FUNCTION_BLOCK VALVE_MANIFOLD (* Migrated from IEC 61131-3 ST *)
  (* Standard: 61499-2 *)
  (* Version 1.0, 2026-11-06, st2fb *)
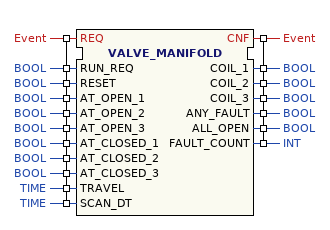
  EVENT_INPUT
    REQ WITH RUN_REQ, RESET, AT_OPEN_1, AT_OPEN_2, AT_OPEN_3, AT_CLOSED_1, AT_CLOSED_2, AT_CLOSED_3, TRAVEL, SCAN_DT;
  END_EVENT
  EVENT_OUTPUT
    CNF WITH COIL_1, COIL_2, COIL_3, ANY_FAULT, ALL_OPEN, FAULT_COUNT;
  END_EVENT
  VAR_INPUT
    RUN_REQ : BOOL;
    RESET : BOOL;
    AT_OPEN_1 : BOOL;
    AT_OPEN_2 : BOOL;
    AT_OPEN_3 : BOOL;
    AT_CLOSED_1 : BOOL;
    AT_CLOSED_2 : BOOL;
    AT_CLOSED_3 : BOOL;
    TRAVEL : TIME;
    SCAN_DT : TIME;
  END_VAR
  VAR_OUTPUT
    COIL_1 : BOOL;
    COIL_2 : BOOL;
    COIL_3 : BOOL;
    ANY_FAULT : BOOL;
    ALL_OPEN : BOOL;
    FAULT_COUNT : INT;
  END_VAR
  VAR
    ST2FB_NOW : TIME := T#0s;
    V1_OPEN_CMD : BOOL;
    V1_COIL : BOOL;
    V1_FAULT : BOOL;
    V1_OPENED : BOOL;
    V1_W_IN : BOOL;
    V1_W_PT : TIME;
    V1_W_Q : BOOL;
    V1_W_ET : TIME;
    V1_W_STATE : INT;
    V1_W_PREV_IN : BOOL;
    V1_W_START_TIME : TIME;
    V2_OPEN_CMD : BOOL;
    V2_COIL : BOOL;
    V2_FAULT : BOOL;
    V2_OPENED : BOOL;
    V2_W_IN : BOOL;
    V2_W_PT : TIME;
    V2_W_Q : BOOL;
    V2_W_ET : TIME;
    V2_W_STATE : INT;
    V2_W_PREV_IN : BOOL;
    V2_W_START_TIME : TIME;
    V3_OPEN_CMD : BOOL;
    V3_COIL : BOOL;
    V3_FAULT : BOOL;
    V3_OPENED : BOOL;
    V3_W_IN : BOOL;
    V3_W_PT : TIME;
    V3_W_Q : BOOL;
    V3_W_ET : TIME;
    V3_W_STATE : INT;
    V3_W_PREV_IN : BOOL;
    V3_W_START_TIME : TIME;
  END_VAR
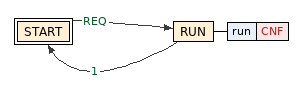
  EC_STATES
    START;
    RUN : run -> CNF;
  END_STATES
  EC_TRANSITIONS
    START TO RUN := REQ;
    RUN TO START := 1;
  END_TRANSITIONS
  ALGORITHM run IN ST:
ST2FB_NOW := ST2FB_NOW + SCAN_DT;

(* V1 *)
V1_OPEN_CMD := RUN_REQ AND NOT ANY_FAULT;
V1_COIL := V1_OPEN_CMD AND NOT V1_FAULT;
V1_W_IN := (V1_COIL AND NOT AT_OPEN_1) OR (NOT V1_COIL AND NOT AT_CLOSED_1 AND NOT V1_FAULT);
V1_W_PT := TRAVEL;
IF (V1_W_STATE = 0) AND NOT V1_W_PREV_IN AND V1_W_IN THEN
  V1_W_STATE := 1;
  V1_W_Q := FALSE;
  V1_W_START_TIME := ST2FB_NOW;
ELSE
  IF NOT V1_W_IN THEN
    V1_W_ET := T#0s;
    V1_W_Q := FALSE;
    V1_W_STATE := 0;
  ELSIF V1_W_STATE = 1 THEN
    IF V1_W_START_TIME + V1_W_PT <= ST2FB_NOW THEN
      V1_W_STATE := 2;
      V1_W_Q := TRUE;
      V1_W_ET := V1_W_PT;
    ELSE
      V1_W_ET := ST2FB_NOW - V1_W_START_TIME;
    END_IF;
  END_IF;
END_IF;
V1_W_PREV_IN := V1_W_IN;
V1_FAULT := V1_W_Q OR (NOT RESET AND V1_FAULT);
V1_OPENED := V1_COIL AND AT_OPEN_1 AND NOT AT_CLOSED_1;

(* V2 *)
V2_OPEN_CMD := V1_OPENED;
V2_COIL := V2_OPEN_CMD AND NOT V2_FAULT;
V2_W_IN := (V2_COIL AND NOT AT_OPEN_2) OR (NOT V2_COIL AND NOT AT_CLOSED_2 AND NOT V2_FAULT);
V2_W_PT := TRAVEL;
IF (V2_W_STATE = 0) AND NOT V2_W_PREV_IN AND V2_W_IN THEN
  V2_W_STATE := 1;
  V2_W_Q := FALSE;
  V2_W_START_TIME := ST2FB_NOW;
ELSE
  IF NOT V2_W_IN THEN
    V2_W_ET := T#0s;
    V2_W_Q := FALSE;
    V2_W_STATE := 0;
  ELSIF V2_W_STATE = 1 THEN
    IF V2_W_START_TIME + V2_W_PT <= ST2FB_NOW THEN
      V2_W_STATE := 2;
      V2_W_Q := TRUE;
      V2_W_ET := V2_W_PT;
    ELSE
      V2_W_ET := ST2FB_NOW - V2_W_START_TIME;
    END_IF;
  END_IF;
END_IF;
V2_W_PREV_IN := V2_W_IN;
V2_FAULT := V2_W_Q OR (NOT RESET AND V2_FAULT);
V2_OPENED := V2_COIL AND AT_OPEN_2 AND NOT AT_CLOSED_2;

(* V3 *)
V3_OPEN_CMD := V2_OPENED;
V3_COIL := V3_OPEN_CMD AND NOT V3_FAULT;
V3_W_IN := (V3_COIL AND NOT AT_OPEN_3) OR (NOT V3_COIL AND NOT AT_CLOSED_3 AND NOT V3_FAULT);
V3_W_PT := TRAVEL;
IF (V3_W_STATE = 0) AND NOT V3_W_PREV_IN AND V3_W_IN THEN
  V3_W_STATE := 1;
  V3_W_Q := FALSE;
  V3_W_START_TIME := ST2FB_NOW;
ELSE
  IF NOT V3_W_IN THEN
    V3_W_ET := T#0s;
    V3_W_Q := FALSE;
    V3_W_STATE := 0;
  ELSIF V3_W_STATE = 1 THEN
    IF V3_W_START_TIME + V3_W_PT <= ST2FB_NOW THEN
      V3_W_STATE := 2;
      V3_W_Q := TRUE;
      V3_W_ET := V3_W_PT;
    ELSE
      V3_W_ET := ST2FB_NOW - V3_W_START_TIME;
    END_IF;
  END_IF;
END_IF;
V3_W_PREV_IN := V3_W_IN;
V3_FAULT := V3_W_Q OR (NOT RESET AND V3_FAULT);
V3_OPENED := V3_COIL AND AT_OPEN_3 AND NOT AT_CLOSED_3;

COIL_1 := V1_COIL;
COIL_2 := V2_COIL;
COIL_3 := V3_COIL;
FAULT_COUNT := 0;
IF V1_FAULT THEN
  FAULT_COUNT := FAULT_COUNT + 1;
END_IF;
IF V2_FAULT THEN
  FAULT_COUNT := FAULT_COUNT + 1;
END_IF;
IF V3_FAULT THEN
  FAULT_COUNT := FAULT_COUNT + 1;
END_IF;
ANY_FAULT := FAULT_COUNT > 0;
ALL_OPEN := V3_OPENED;
  END_ALGORITHM
END_FUNCTION_BLOCK
